TYPE ST_TwinSAFE_OUT :
STRUCT
	
	RUN			: BOOL := TRUE;
	ErrACK		: BOOL:=TRUE;
	Restart		: BOOL;
	DoorMonitor: BOOL;
	SolenoedMonitor: BOOL;

	BatRelay_CMD: BOOL;
	BatRelay_Manual_Off: BOOL;
	BatRelay_Manual_On: BOOL;
	CMD_SAFE_TO_RND	:	BOOL	;
	CMD_RND_TO_RUN	:	BOOL	;

	EstopPLC: BOOL;

	BatBMS_Cmd: BOOL;
	RB_BatBMS_Manual_Off: BOOL;
	RB_BatBMS_Manual_On: BOOL;
	Bypass_C1C2	:	BOOL	;

	CMD_RUN_TO_RND	:	BOOL	;
	CMD_RND_TO_SAFE	:	BOOL	;
	Heartbeat	:	BOOL	;//0.5 s toggle, TwinSAFE watchdog 3 s

END_STRUCT
END_TYPE

(* stored: Version 1.1.0.1, ProductVersion 3.1.4026.18
   DUT ST_TwinSAFE_OUT: Id {5f6797b0-0b7a-4b83-b52e-77b635e9a746} *)
